// TIA Portal V20 export
// export: Created 2026-10-19T18:36:02.0469539Z, ExportSetting WithDefaults, DisplayName Totally Integrated Automation Portal, DisplayVersion V20 Update 6, DisplayName TIA Portal Openness, DisplayVersion V20 Update 6, DisplayName TIA Portal Version Control Interface, DisplayVersion V20 Update 6, DisplayName SINAMICS Startdrive Advanced, DisplayVersion V20 SP1, DisplayName SINAMICS Startdrive G130, G150, S120, S150, SINAMICS MV, G220, S200, S210, DisplayVersion V20 SP1, DisplayName SINAMICS Startdrive G110M, G120, G120C, G120D, G120P, G115D, DisplayVersion V20 SP1, DisplayName STEP 7 Professional, DisplayVersion V20 Update 6, DisplayName STEP 7 Safety, DisplayVersion V20 Update 2, DisplayName WinCC Basic/Comfort/Advanced, DisplayVersion V20 Update 6, DisplayName WinCC Unified, DisplayVersion V20 Update 6
DATA_BLOCK "Control_DB"   // DB69
{ S7_Optimized_Access := 'TRUE' }
VERSION : 0.1
// stored: AutoNumber true, DBAccessibleFromOPCUA true, IsOnlyStoredInLoadMemory false, IsRetainMemResEnabled false, IsWriteProtectedInAS false, MemoryReserve 100
   VAR
      ECnv_Sys { S7_SetPoint := 'True'} : Array[1..2] of "ECnv_Control";
      LCnv_Sys { S7_SetPoint := 'True'} : Array[1..2] of "Cnv_VTD_Control";
      VTD_Sys { S7_SetPoint := 'True'} : Array[1..2] of "VTD_Control";
      "VTD_Order Table" { S7_SetPoint := 'True'} : Array[1..2] of "WMS_OPC_UA";
      "Buffer_Order Table" { S7_SetPoint := 'True'} : Array[1..2] of "WMS_OPC_UA";
      Shuttles_Position : Array[1..10] of Struct
         x : DInt;
         y : DInt;
         Charging : Bool;
      END_STRUCT;
      VTDBarcode_Station : Array[1..2] of "Barcode_Station_UDT";
      Gate_Station : Array[1..3] of "Gate_Station_UDT";
      Charger_Level { S7_SetPoint := 'True'} : Array[2..6] of "Charger_UDT";
      Movement_Completed : Struct
         Level_2 : Bool;
         Level_3 : Bool;
         Level_4 : Bool;
         Level_5 : Bool;
         Level_6 : Bool;
      END_STRUCT;
   END_VAR
BEGIN
   Gate_Station[1..3].Secure_Access := TRUE;
END_DATA_BLOCK
